(* Logix 5000 project; controller NWGG_Treater_Dayton vendor 1 type 14 code 238 rev 35.11; software revision 35.00; part 2 of 5 *)

ADD_ON_INSTRUCTION SAI_CheckAlive   (* revision 1.0, vendor Jimmy Gao *)
VAR_INPUT
   HeartBeat : BOOL; {required}
END_VAR
VAR_OUTPUT
   Alive : BOOL; {access Read Only, visible}
END_VAR
VAR
   bResetTimer : BOOL; {access None}
   ons : DINT; {access None}
   TON : TIMER; {access None}
END_VAR

ROUTINE Logic   (* ladder *)
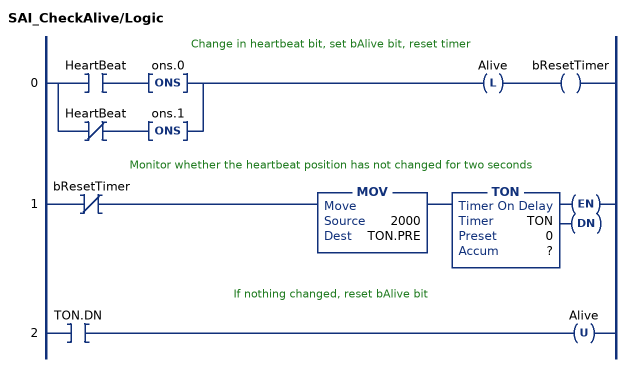
   // Change in heartbeat bit, set bAlive bit, reset timer
   0: [XIC(HeartBeat) ONS(ons.0) ,XIO(HeartBeat) ONS(ons.1) ]OTL(Alive)OTE(bResetTimer);
   // Monitor whether the heartbeat position has not changed for two seconds
   1: XIO(bResetTimer)MOV(2000,TON.PRE)TON(TON,?,?);
   // If nothing changed, reset bAlive bit
   2: XIC(TON.DN)OTU(Alive);
END_ROUTINE
END_ADD_ON_INSTRUCTION

ADD_ON_INSTRUCTION SAI_IND_CalFree   (* revision 1.0, vendor Griffin Hodnett *)
VAR_INPUT
   RatedCapacity : REAL; {required}
   ScaleUnit : DINT; {required}
   RatedOutput : REAL; {access None, required}
   Start : BOOL; {visible}
END_VAR
VAR_OUTPUT
   Done : BOOL; {access Read Only, visible}
   Error : BOOL; {access Read Only, visible}
   Status : DINT; {access Read Only, visible}
END_VAR
VAR_IN_OUT
   MSG_CalFreeTrigger : MESSAGE; {required}
   MSG_CalFreeStatus : MESSAGE; {required}
   MSG_CalFreeUnit : MESSAGE; {required}
   MSG_CalFreeCellCapacity : MESSAGE; {required}
   MSG_CalFreeCellOutput : MESSAGE; {required}
   TmpTrigger : INT; {required}
   TmpAdjStatus : INT; {required}
END_VAR
VAR
   ons : DINT; {access None}
   Step : INT; {access None}
   TON : TIMER[7]; {access None}
   EnterAdj : BOOL; {access None}
   EnterCancel : BOOL; {access None}
END_VAR

ROUTINE Logic   (* ladder *)
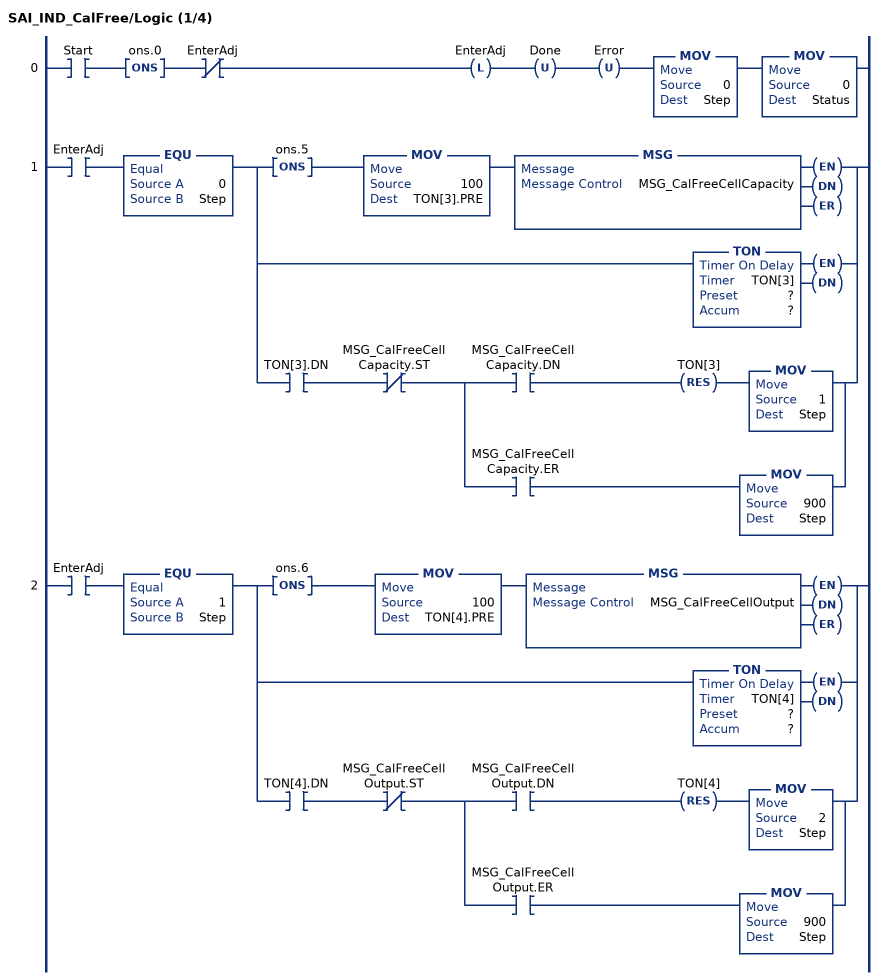
   0: XIC(Start)ONS(ons.0)XIO(EnterAdj)OTL(EnterAdj)OTU(Done)OTU(Error)MOV(0,Step)MOV(0,Status);
   1: XIC(EnterAdj)EQU(0,Step)[[ONS(ons.5) MOV(100,TON[3].PRE) MSG(MSG_CalFreeCellCapacity) ,TON(TON[3],?,?) ] ,XIC(TON[3].DN) XIO(MSG_CalFreeCellCapacity.ST) [XIC(MSG_CalFreeCellCapacity.DN) RES(TON[3]) MOV(1,Step) ,XIC(MSG_CalFreeCellCapacity.ER) MOV(900,Step) ] ];
   2: XIC(EnterAdj)EQU(1,Step)[[ONS(ons.6) MOV(100,TON[4].PRE) MSG(MSG_CalFreeCellOutput) ,TON(TON[4],?,?) ] ,XIC(TON[4].DN) XIO(MSG_CalFreeCellOutput.ST) [XIC(MSG_CalFreeCellOutput.DN) RES(TON[4]) MOV(2,Step) ,XIC(MSG_CalFreeCellOutput.ER) MOV(900,Step) ] ];
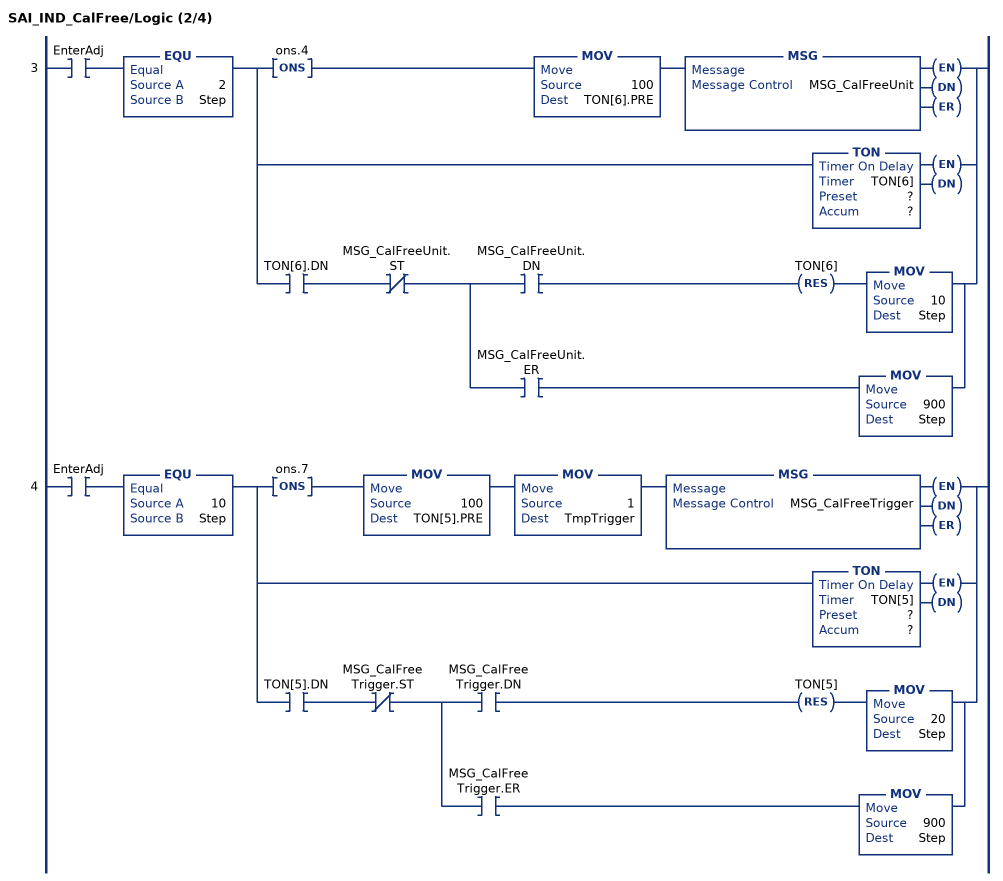
   3: XIC(EnterAdj)EQU(2,Step)[[ONS(ons.4) MOV(100,TON[6].PRE) MSG(MSG_CalFreeUnit) ,TON(TON[6],?,?) ] ,XIC(TON[6].DN) XIO(MSG_CalFreeUnit.ST) [XIC(MSG_CalFreeUnit.DN) RES(TON[6]) MOV(10,Step) ,XIC(MSG_CalFreeUnit.ER) MOV(900,Step) ] ];
   4: XIC(EnterAdj)EQU(10,Step)[[ONS(ons.7) MOV(100,TON[5].PRE) MOV(1,TmpTrigger) MSG(MSG_CalFreeTrigger) ,TON(TON[5],?,?) ] ,XIC(TON[5].DN) XIO(MSG_CalFreeTrigger.ST) [XIC(MSG_CalFreeTrigger.DN) RES(TON[5]) MOV(20,Step) ,XIC(MSG_CalFreeTrigger.ER) MOV(900,Step) ] ];
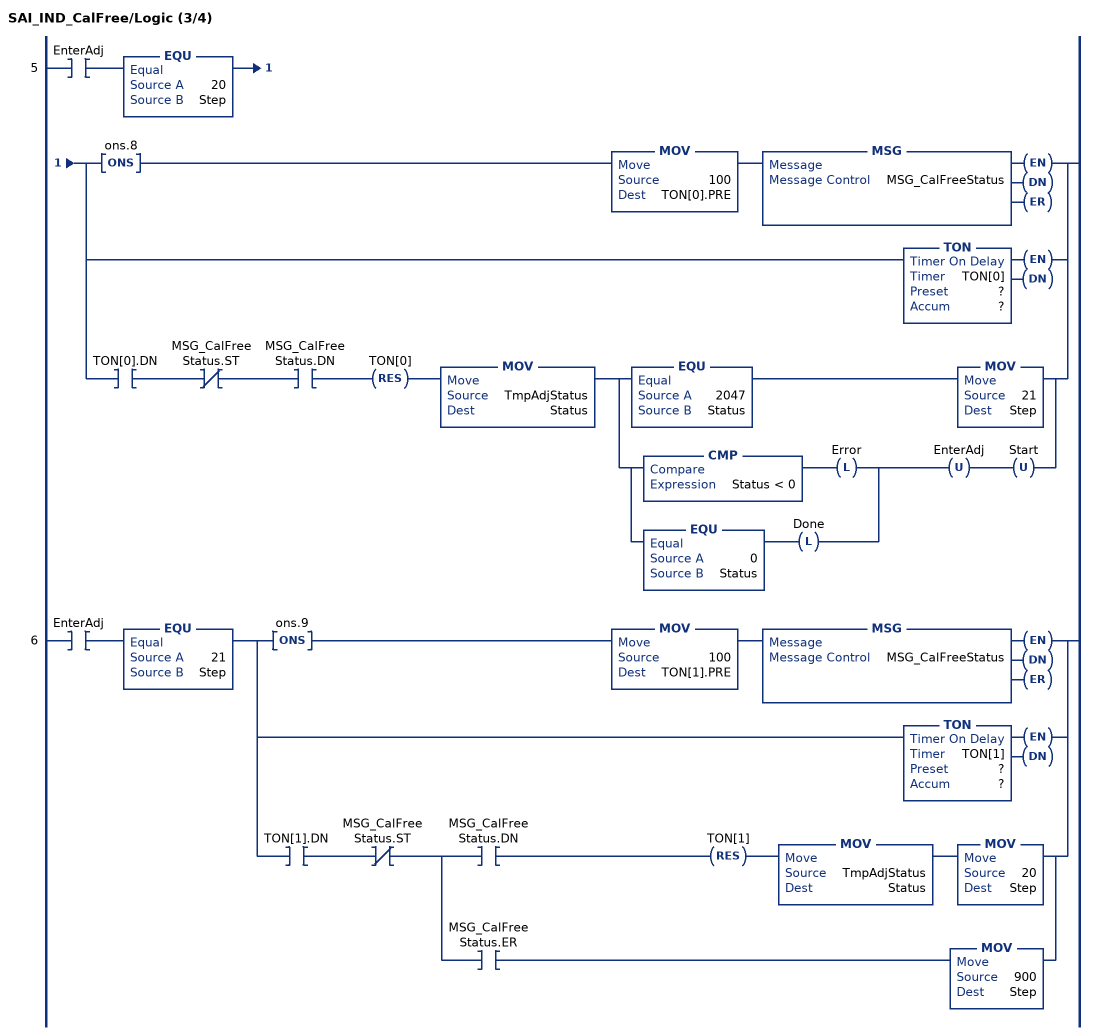
   5: XIC(EnterAdj)EQU(20,Step)[[ONS(ons.8) MOV(100,TON[0].PRE) MSG(MSG_CalFreeStatus) ,TON(TON[0],?,?) ] ,XIC(TON[0].DN) XIO(MSG_CalFreeStatus.ST) XIC(MSG_CalFreeStatus.DN) RES(TON[0]) MOV(TmpAdjStatus,Status) [EQU(2047,Status) MOV(21,Step) ,[CMP(Status < 0) OTL(Error) ,EQU(0,Status) OTL(Done) ] OTU(EnterAdj) OTU(Start) ] ];
   6: XIC(EnterAdj)EQU(21,Step)[[ONS(ons.9) MOV(100,TON[1].PRE) MSG(MSG_CalFreeStatus) ,TON(TON[1],?,?) ] ,XIC(TON[1].DN) XIO(MSG_CalFreeStatus.ST) [XIC(MSG_CalFreeStatus.DN) RES(TON[1]) MOV(TmpAdjStatus,Status) MOV(20,Step) ,XIC(MSG_CalFreeStatus.ER) MOV(900,Step) ] ];
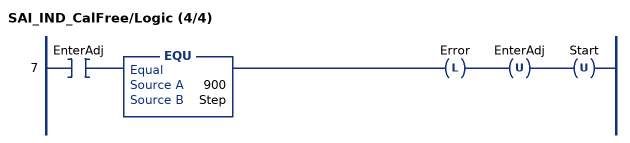
   7: XIC(EnterAdj)EQU(900,Step)OTL(Error)OTU(EnterAdj)OTU(Start);
END_ROUTINE
END_ADD_ON_INSTRUCTION

ADD_ON_INSTRUCTION SAI_IND_ReadAdjustSettings   (* revision 1.0, vendor Griffin Hodnett *)
VAR_INPUT
   Read : BOOL; {visible}
END_VAR
VAR_OUTPUT
   ScaleCapacity : REAL; {visible}
   Increment : REAL; {visible}
   Done : BOOL; {access Read Only, visible}
   Error : BOOL; {access Read Only, visible}
END_VAR
VAR_IN_OUT
   MSG_ReadCap : MESSAGE; {required}
   MSG_ReadInc : MESSAGE; {required}
   TmpInc : REAL; {required}
   TmpCapacity : REAL; {required}
END_VAR
VAR
   TON : TIMER[1]; {access None}
   Step : INT; {access None}
   Get_Values : BOOL; {access None}
   ons : DINT; {access None}
END_VAR

ROUTINE Logic   (* ladder *)
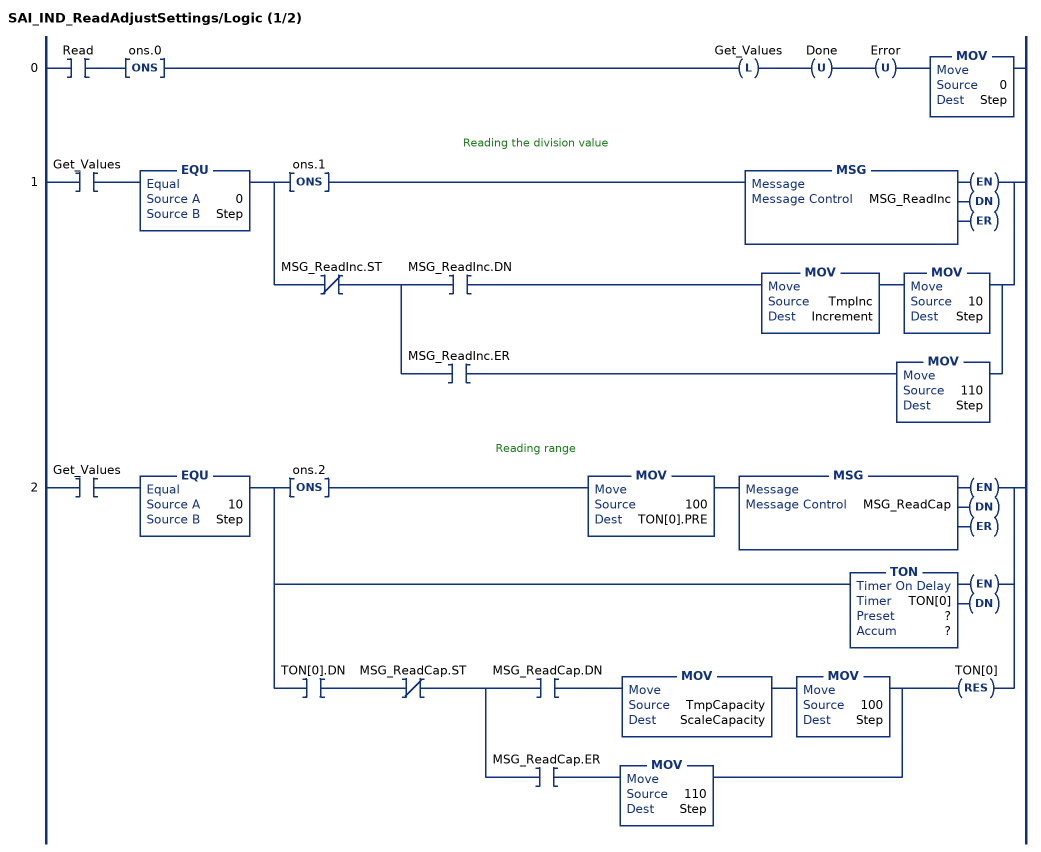
   0: XIC(Read)ONS(ons.0)OTL(Get_Values)OTU(Done)OTU(Error)MOV(0,Step);
   // Reading the division value
   1: XIC(Get_Values)EQU(0,Step)[ONS(ons.1) MSG(MSG_ReadInc) ,XIO(MSG_ReadInc.ST) [XIC(MSG_ReadInc.DN) MOV(TmpInc,Increment) MOV(10,Step) ,XIC(MSG_ReadInc.ER) MOV(110,Step) ] ];
   // Reading range
   2: XIC(Get_Values)EQU(10,Step)[[ONS(ons.2) MOV(100,TON[0].PRE) MSG(MSG_ReadCap) ,TON(TON[0],?,?) ] ,XIC(TON[0].DN) XIO(MSG_ReadCap.ST) [XIC(MSG_ReadCap.DN) MOV(TmpCapacity,ScaleCapacity) MOV(100,Step) ,XIC(MSG_ReadCap.ER) MOV(110,Step) ] RES(TON[0]) ];
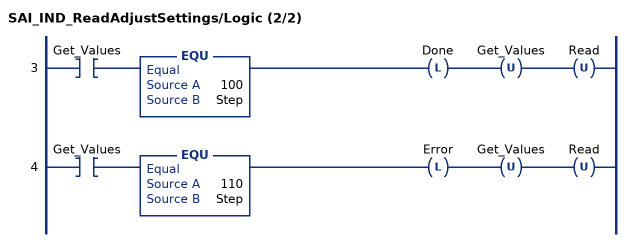
   3: XIC(Get_Values)EQU(100,Step)OTL(Done)OTU(Get_Values)OTU(Read);
   4: XIC(Get_Values)EQU(110,Step)OTL(Error)OTU(Get_Values)OTU(Read);
END_ROUTINE
END_ADD_ON_INSTRUCTION

ADD_ON_INSTRUCTION SAI_IND_SpanAdjust   (* revision 1.0, vendor Griffin Hodnett *)
VAR_INPUT
   LinearityRange : INT; {access None, required}
   Hi_Weight : REAL; {visible}
   Mid_Weight : REAL; {visible}
   Low_Weight : REAL; {visible}
   xLow_Weight : REAL; {visible}
   Start : BOOL; {visible}
END_VAR
VAR_OUTPUT
   CurrentWeight : REAL; {access Read Only, visible}
END_VAR
VAR_INPUT
   ConfirmWeight : BOOL; {visible}
   Cancel : BOOL; {visible}
END_VAR
VAR_OUTPUT
   Done : BOOL; {access Read Only, visible}
   Error : BOOL; {access Read Only, visible}
   Cancelled : BOOL; {access Read Only, visible}
   LoadWeight : BOOL; {access Read Only, visible}
END_VAR
VAR_INPUT
   DataOK : BOOL; {required}
END_VAR
VAR_OUTPUT
   Status : INT; {access Read Only, visible}
   CurrentPoint : DINT; {access Read Only, visible}
END_VAR
VAR_IN_OUT
   MSG_CancelAdj : MESSAGE; {required}
   MSG_StartSpanAdj : MESSAGE; {required}
   MSG_LinearityRange : MESSAGE; {required}
   MSG_ReadAdjStatus : MESSAGE; {required}
   MSG_ValidateAdj : MESSAGE; {required}
   TmpTrigger : SINT; {required}
   TmpAdjStatus : INT; {required}
   TmpSpanAdjWeight : REAL; {required}
END_VAR
VAR
   Step : INT; {access None}
   TON : TIMER[3]; {access None}
   ons : DINT; {access None}
   EnterCancel : BOOL; {access None}
   EnterAdj : BOOL; {access None}
   WeightCheck : BOOL; {access None}
END_VAR

ROUTINE Logic   (* ladder *)
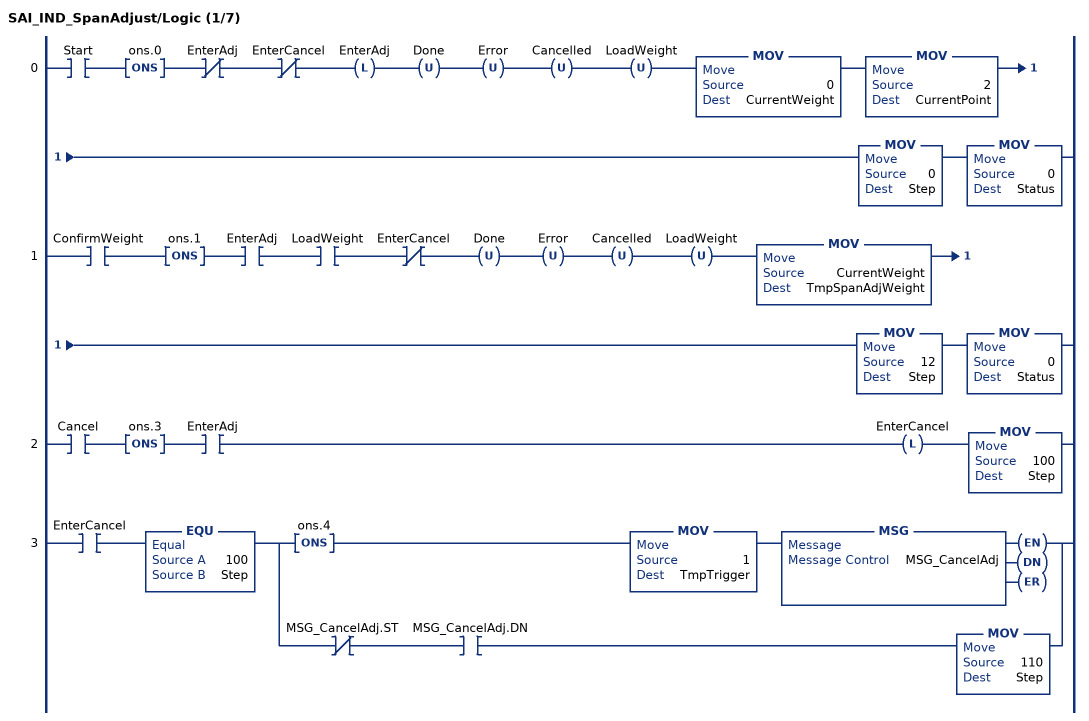
   0: XIC(Start)ONS(ons.0)XIO(EnterAdj)XIO(EnterCancel)OTL(EnterAdj)OTU(Done)OTU(Error)OTU(Cancelled)OTU(LoadWeight)MOV(0,CurrentWeight)MOV(2,CurrentPoint)MOV(0,Step)MOV(0,Status);
   1: XIC(ConfirmWeight)ONS(ons.1)XIC(EnterAdj)XIC(LoadWeight)XIO(EnterCancel)OTU(Done)OTU(Error)OTU(Cancelled)OTU(LoadWeight)MOV(CurrentWeight,TmpSpanAdjWeight)MOV(12,Step)MOV(0,Status);
   2: XIC(Cancel)ONS(ons.3)XIC(EnterAdj)OTL(EnterCancel)MOV(100,Step);
   3: XIC(EnterCancel)EQU(100,Step)[ONS(ons.4) MOV(1,TmpTrigger) MSG(MSG_CancelAdj) ,XIO(MSG_CancelAdj.ST) XIC(MSG_CancelAdj.DN) MOV(110,Step) ];
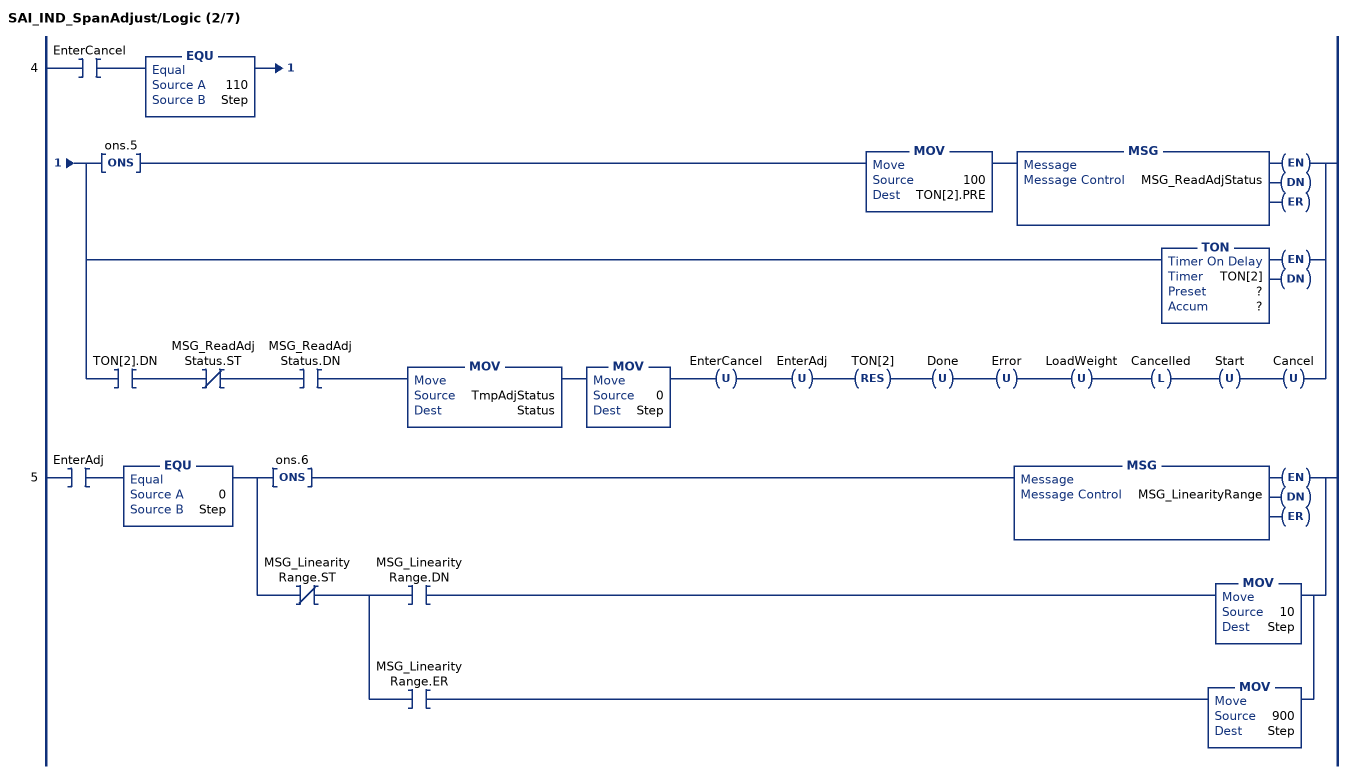
   4: XIC(EnterCancel)EQU(110,Step)[[ONS(ons.5) MOV(100,TON[2].PRE) MSG(MSG_ReadAdjStatus) ,TON(TON[2],?,?) ] ,XIC(TON[2].DN) XIO(MSG_ReadAdjStatus.ST) XIC(MSG_ReadAdjStatus.DN) MOV(TmpAdjStatus,Status) MOV(0,Step) OTU(EnterCancel) OTU(EnterAdj) RES(TON[2]) OTU(Done) OTU(Error) OTU(LoadWeight) OTL(Cancelled) OTU(Start) OTU(Cancel) ];
   5: XIC(EnterAdj)EQU(0,Step)[ONS(ons.6) MSG(MSG_LinearityRange) ,XIO(MSG_LinearityRange.ST) [XIC(MSG_LinearityRange.DN) MOV(10,Step) ,XIC(MSG_LinearityRange.ER) MOV(900,Step) ] ];
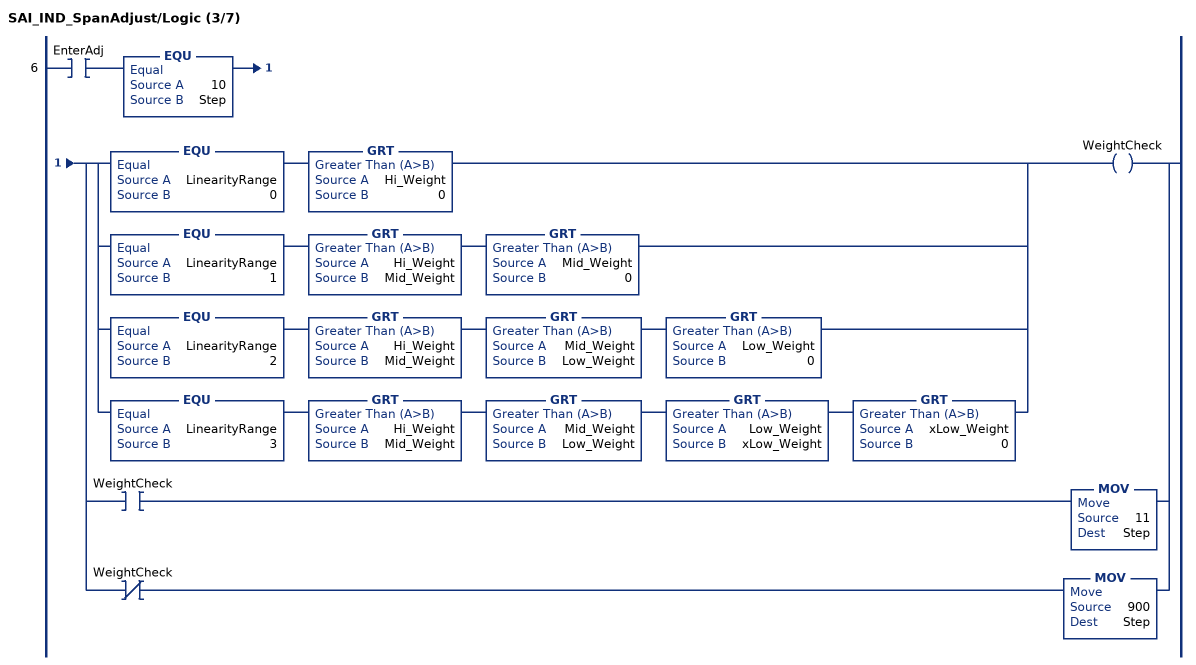
   6: XIC(EnterAdj)EQU(10,Step)[[EQU(LinearityRange,0) GRT(Hi_Weight,0) ,[EQU(LinearityRange,1) GRT(Hi_Weight,Mid_Weight) GRT(Mid_Weight,0) ,[EQU(LinearityRange,2) GRT(Hi_Weight,Mid_Weight) GRT(Mid_Weight,Low_Weight) GRT(Low_Weight,0) ,EQU(LinearityRange,3) GRT(Hi_Weight,Mid_Weight) GRT(Mid_Weight,Low_Weight) GRT(Low_Weight,xLow_Weight) GRT(xLow_Weight,0) ] ] ] OTE(WeightCheck) ,[XIC(WeightCheck) MOV(11,Step) ,XIO(WeightCheck) MOV(900,Step) ] ];
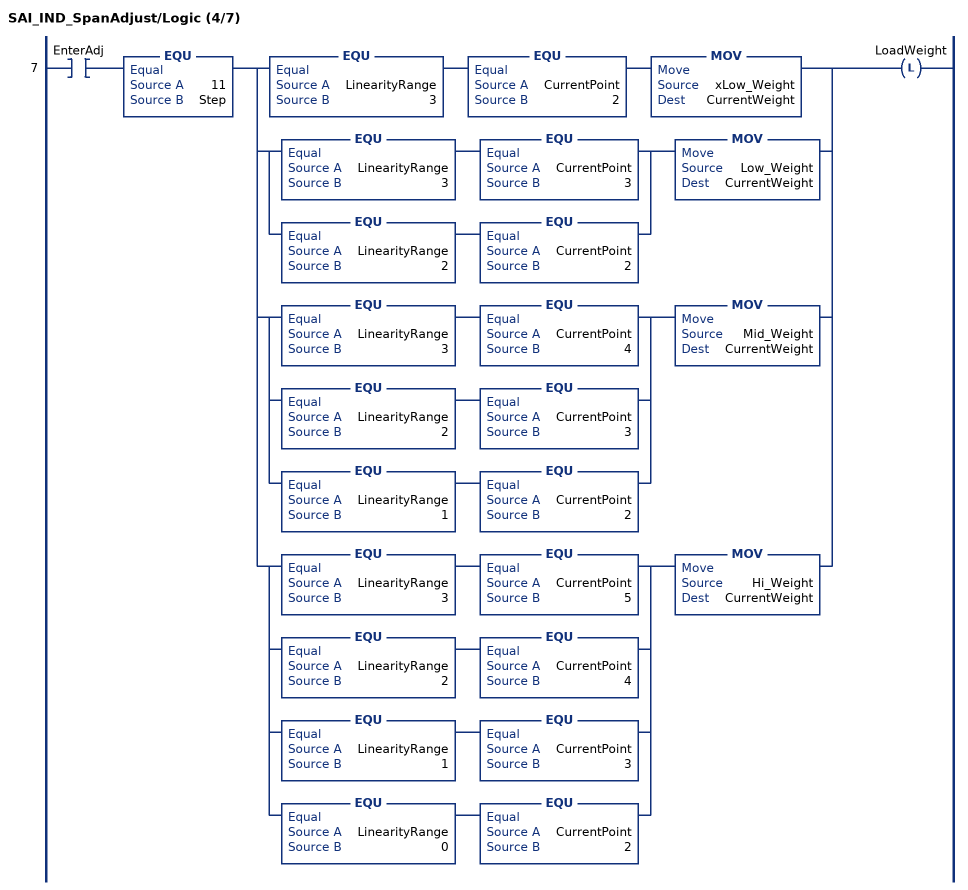
   7: XIC(EnterAdj)EQU(11,Step)[EQU(LinearityRange,3) EQU(CurrentPoint,2) MOV(xLow_Weight,CurrentWeight) ,[[[EQU(LinearityRange,3) EQU(CurrentPoint,3) ,EQU(LinearityRange,2) EQU(CurrentPoint,2) ] MOV(Low_Weight,CurrentWeight) ,[EQU(LinearityRange,3) EQU(CurrentPoint,4) ,[EQU(LinearityRange,2) EQU(CurrentPoint,3) ,EQU(LinearityRange,1) EQU(CurrentPoint,2) ] ] MOV(Mid_Weight,CurrentWeight) ] ,[EQU(LinearityRange,3) EQU(CurrentPoint,5) ,[EQU(LinearityRange,2) EQU(CurrentPoint,4) ,[EQU(LinearityRange,1) EQU(CurrentPoint,3) ,EQU(LinearityRange,0) EQU(CurrentPoint,2) ] ] ] MOV(Hi_Weight,CurrentWeight) ] ]OTL(LoadWeight);
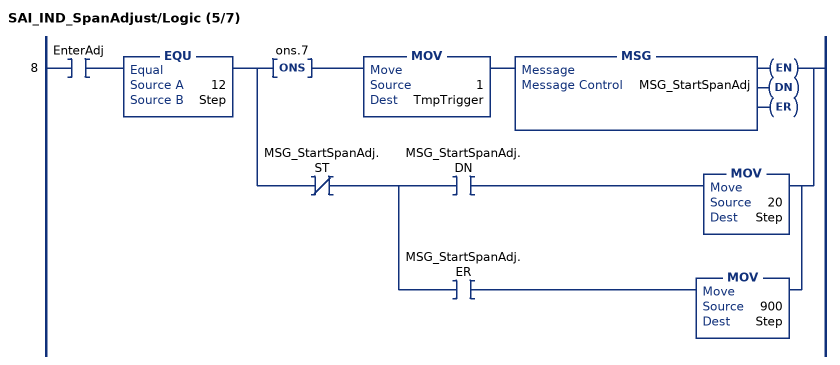
   8: XIC(EnterAdj)EQU(12,Step)[ONS(ons.7) MOV(1,TmpTrigger) MSG(MSG_StartSpanAdj) ,XIO(MSG_StartSpanAdj.ST) [XIC(MSG_StartSpanAdj.DN) MOV(20,Step) ,XIC(MSG_StartSpanAdj.ER) MOV(900,Step) ] ];
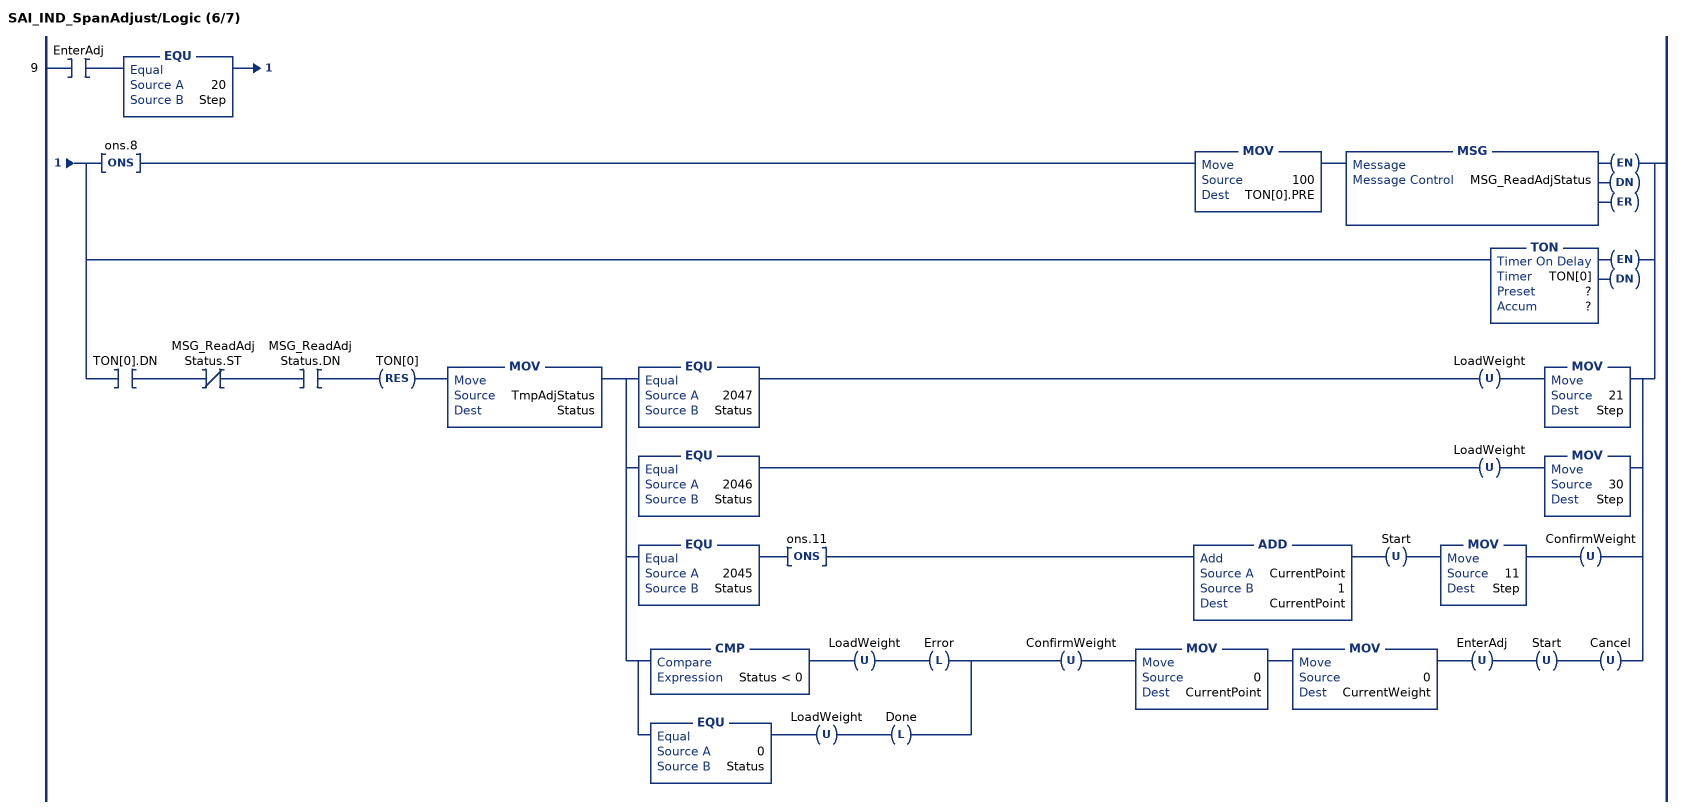
   9: XIC(EnterAdj)EQU(20,Step)[[ONS(ons.8) MOV(100,TON[0].PRE) MSG(MSG_ReadAdjStatus) ,TON(TON[0],?,?) ] ,XIC(TON[0].DN) XIO(MSG_ReadAdjStatus.ST) XIC(MSG_ReadAdjStatus.DN) RES(TON[0]) MOV(TmpAdjStatus,Status) [EQU(2047,Status) OTU(LoadWeight) MOV(21,Step) ,[[EQU(2046,Status) OTU(LoadWeight) MOV(30,Step) ,EQU(2045,Status) ONS(ons.11) ADD(CurrentPoint,1,CurrentPoint) OTU(Start) MOV(11,Step) OTU(ConfirmWeight) ] ,[CMP(Status < 0) OTU(LoadWeight) OTL(Error) ,EQU(0,Status) OTU(LoadWeight) OTL(Done) ] OTU(ConfirmWeight) MOV(0,CurrentPoint) MOV(0,CurrentWeight) OTU(EnterAdj) OTU(Start) OTU(Cancel) ] ] ];
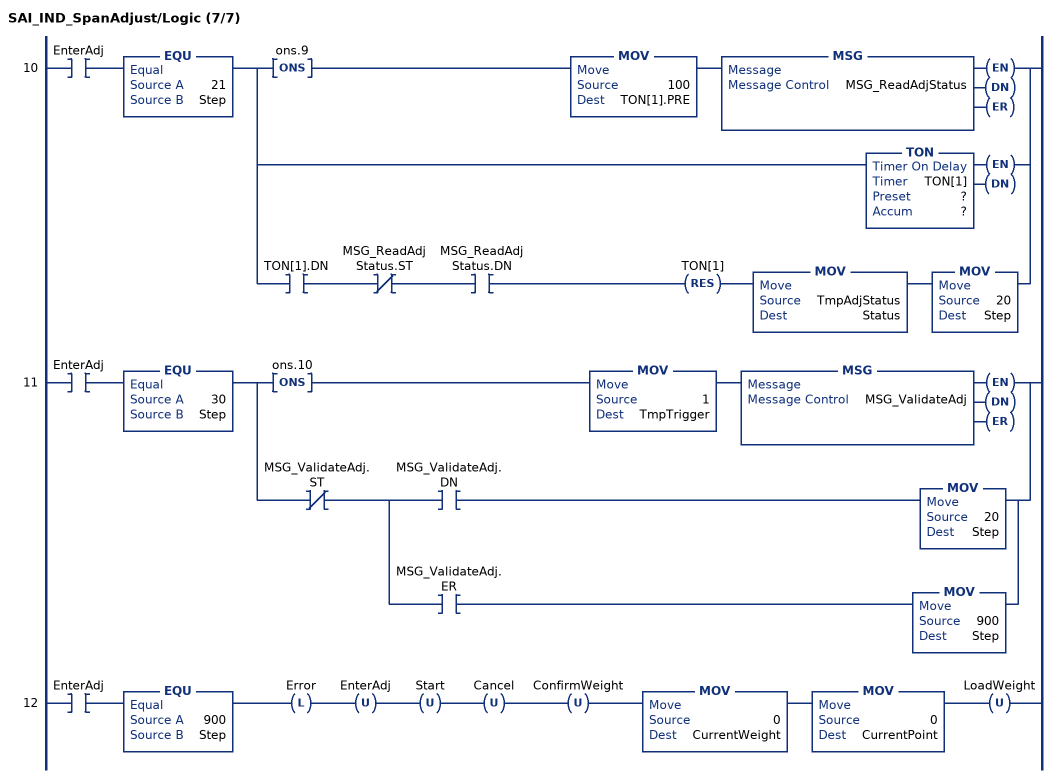
   10: XIC(EnterAdj)EQU(21,Step)[[ONS(ons.9) MOV(100,TON[1].PRE) MSG(MSG_ReadAdjStatus) ,TON(TON[1],?,?) ] ,XIC(TON[1].DN) XIO(MSG_ReadAdjStatus.ST) XIC(MSG_ReadAdjStatus.DN) RES(TON[1]) MOV(TmpAdjStatus,Status) MOV(20,Step) ];
   11: XIC(EnterAdj)EQU(30,Step)[ONS(ons.10) MOV(1,TmpTrigger) MSG(MSG_ValidateAdj) ,XIO(MSG_ValidateAdj.ST) [XIC(MSG_ValidateAdj.DN) MOV(20,Step) ,XIC(MSG_ValidateAdj.ER) MOV(900,Step) ] ];
   12: XIC(EnterAdj)EQU(900,Step)OTL(Error)OTU(EnterAdj)OTU(Start)OTU(Cancel)OTU(ConfirmWeight)MOV(0,CurrentWeight)MOV(0,CurrentPoint)OTU(LoadWeight);
END_ROUTINE
END_ADD_ON_INSTRUCTION

ADD_ON_INSTRUCTION SAI_IND_WeightProc   (* revision 1.0, vendor Griffin Hodnett *)
VAR_INPUT
   WeightCmd : INT; {visible}
   TareImmediate : BOOL; {visible}
   TareStable : BOOL; {visible}
   ZeroImmediate : BOOL; {visible}
   ZeroStable : BOOL; {visible}
   PreTareValue : REAL; {visible}
   PreTare : BOOL; {visible}
   ClearTare : BOOL; {visible}
   MB_Value : REAL; {access Read Only, required}
   MB_Response : INT; {access Read Only, required}
END_VAR
VAR_IN_OUT
   MB_CmdValue : REAL; {required}
END_VAR
VAR_OUTPUT
   MB_Command : INT; {access Read Only, required}
END_VAR
VAR_INPUT
   DataOK : BOOL; {access Read Only, required}
   Motion : BOOL; {access Read Only, required}
   NetMode : BOOL; {required}
   Alarm : BOOL; {required}
END_VAR
VAR_OUTPUT
   RealTimeWeight : REAL; {access Read Only, visible}
   StableWeight : REAL; {access Read Only, visible}
   Done : BOOL; {access Read Only, visible}
   Error : BOOL; {access Read Only, visible}
END_VAR
VAR
   WriteTrigger : BOOL; {access None}
   RestoreTrigger : BOOL; {access None}
   Command : INT; {access None}
   ons : DINT; {access None}
   Prev_WeightCmd : DINT; {access None}
END_VAR

ROUTINE Logic   (* ladder *)
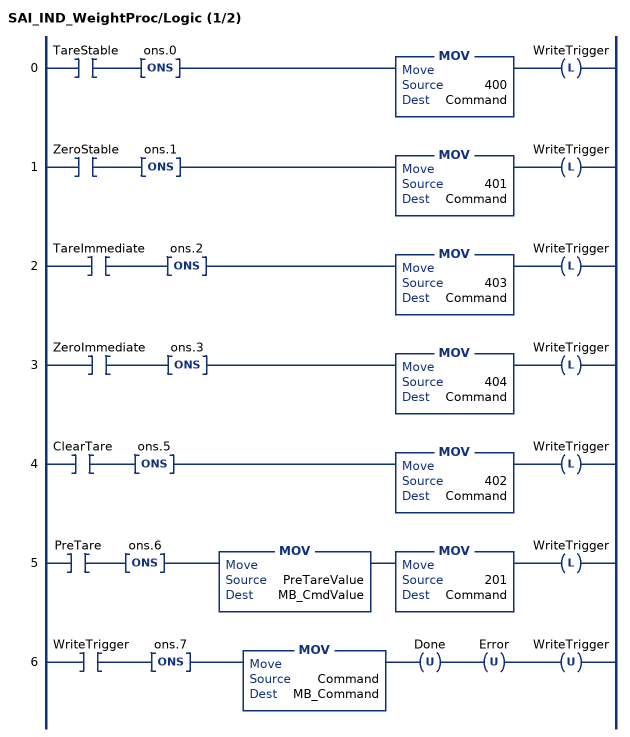
   0: XIC(TareStable)ONS(ons.0)MOV(400,Command)OTL(WriteTrigger);
   1: XIC(ZeroStable)ONS(ons.1)MOV(401,Command)OTL(WriteTrigger);
   2: XIC(TareImmediate)ONS(ons.2)MOV(403,Command)OTL(WriteTrigger);
   3: XIC(ZeroImmediate)ONS(ons.3)MOV(404,Command)OTL(WriteTrigger);
   4: XIC(ClearTare)ONS(ons.5)MOV(402,Command)OTL(WriteTrigger);
   5: XIC(PreTare)ONS(ons.6)MOV(PreTareValue,MB_CmdValue)MOV(201,Command)OTL(WriteTrigger);
   6: XIC(WriteTrigger)ONS(ons.7)MOV(Command,MB_Command)OTU(Done)OTU(Error)OTU(WriteTrigger);
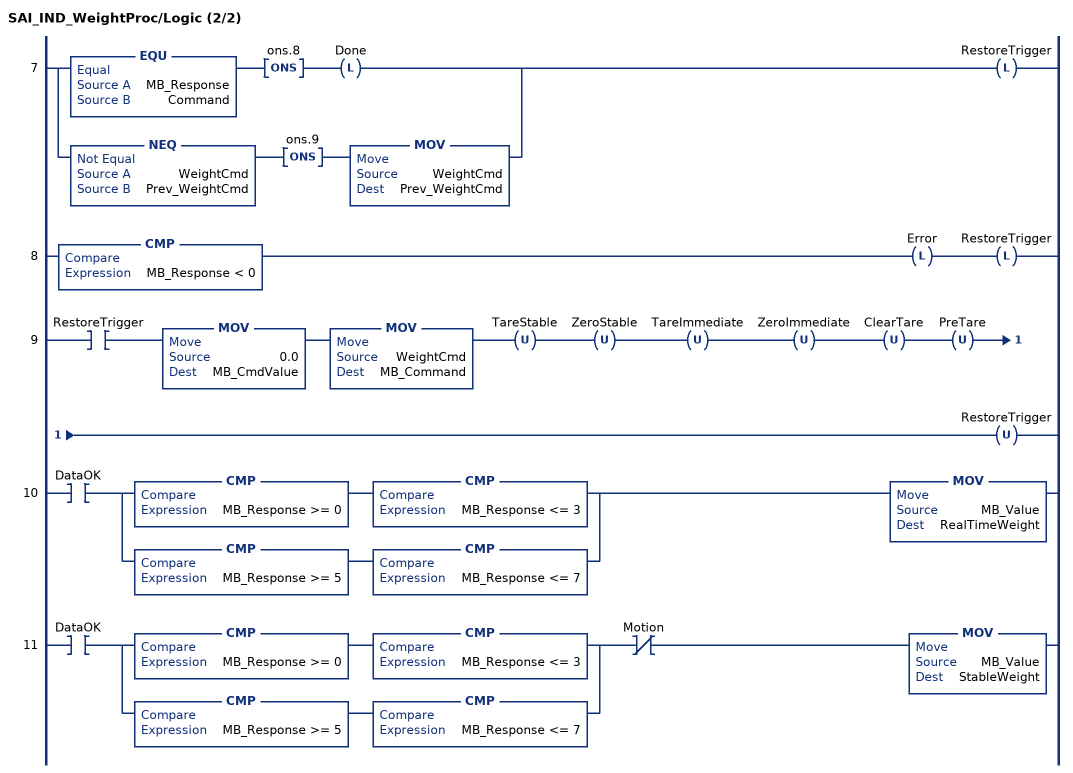
   7: [EQU(MB_Response,Command) ONS(ons.8) OTL(Done) ,NEQ(WeightCmd,Prev_WeightCmd) ONS(ons.9) MOV(WeightCmd,Prev_WeightCmd) ]OTL(RestoreTrigger);
   8: CMP(MB_Response < 0)OTL(Error)OTL(RestoreTrigger);
   9: XIC(RestoreTrigger)MOV(0.0,MB_CmdValue)MOV(WeightCmd,MB_Command)OTU(TareStable)OTU(ZeroStable)OTU(TareImmediate)OTU(ZeroImmediate)OTU(ClearTare)OTU(PreTare)OTU(RestoreTrigger);
   10: XIC(DataOK)[CMP(MB_Response >= 0) CMP(MB_Response <= 3) ,CMP(MB_Response >= 5) CMP(MB_Response <= 7) ]MOV(MB_Value,RealTimeWeight);
   11: XIC(DataOK)[CMP(MB_Response >= 0) CMP(MB_Response <= 3) ,CMP(MB_Response >= 5) CMP(MB_Response <= 7) ]XIO(Motion)MOV(MB_Value,StableWeight);
END_ROUTINE
END_ADD_ON_INSTRUCTION

ADD_ON_INSTRUCTION SAI_IND_WriteAdjustSettings   (* revision 1.0, vendor Griffin Hodnett *)
VAR_INPUT
   ScaleCapacity : REAL; {required}
   Increment : REAL; {required}
   Write : BOOL; {visible}
END_VAR
VAR_OUTPUT
   Done : BOOL; {access Read Only, visible}
   Error : BOOL; {access Read Only, visible}
END_VAR
VAR_IN_OUT
   MSG_WriteCap : MESSAGE; {required}
   MSG_WriteInc : MESSAGE; {required}
END_VAR
VAR
   ons : DINT; {access None}
   Step : INT; {access None}
   TON : TIMER[2]; {access None}
   Write_Values : BOOL; {access None}
END_VAR

ROUTINE Logic   (* ladder *)
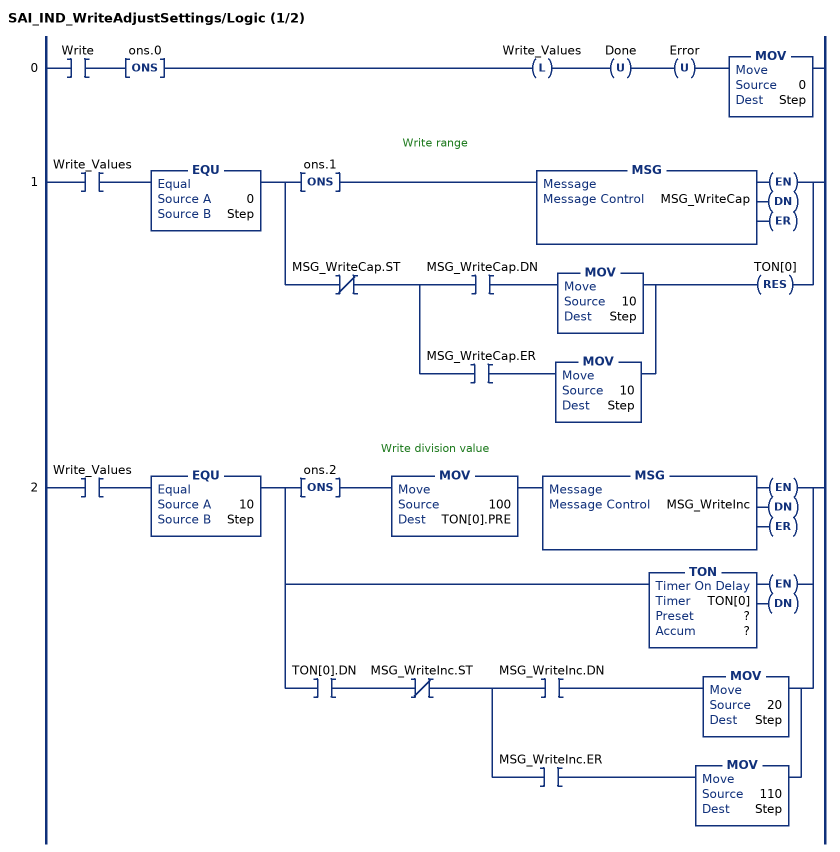
   0: XIC(Write)ONS(ons.0)OTL(Write_Values)OTU(Done)OTU(Error)MOV(0,Step);
   // Write range
   1: XIC(Write_Values)EQU(0,Step)[ONS(ons.1) MSG(MSG_WriteCap) ,XIO(MSG_WriteCap.ST) [XIC(MSG_WriteCap.DN) MOV(10,Step) ,XIC(MSG_WriteCap.ER) MOV(10,Step) ] RES(TON[0]) ];
   // Write division value
   2: XIC(Write_Values)EQU(10,Step)[[ONS(ons.2) MOV(100,TON[0].PRE) MSG(MSG_WriteInc) ,TON(TON[0],?,?) ] ,XIC(TON[0].DN) XIO(MSG_WriteInc.ST) [XIC(MSG_WriteInc.DN) MOV(20,Step) ,XIC(MSG_WriteInc.ER) MOV(110,Step) ] ];
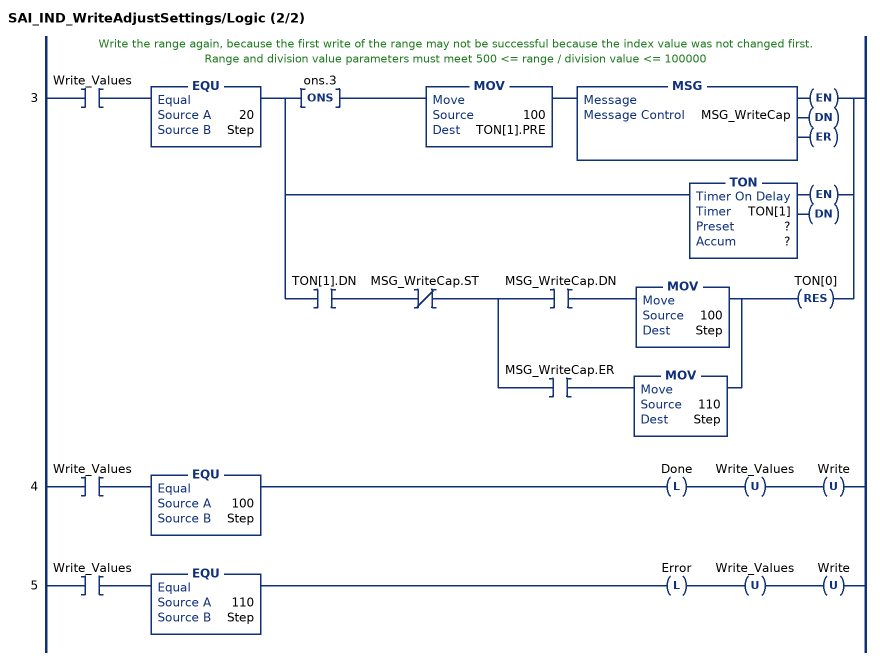
   // Write the range again, because the first write of the range may not be successful because the index value was not changed first.
   // Range and division value parameters must meet 500 <= range / division value <= 100000
   3: XIC(Write_Values)EQU(20,Step)[[ONS(ons.3) MOV(100,TON[1].PRE) MSG(MSG_WriteCap) ,TON(TON[1],?,?) ] ,XIC(TON[1].DN) XIO(MSG_WriteCap.ST) [XIC(MSG_WriteCap.DN) MOV(100,Step) ,XIC(MSG_WriteCap.ER) MOV(110,Step) ] RES(TON[0]) ];
   4: XIC(Write_Values)EQU(100,Step)OTL(Done)OTU(Write_Values)OTU(Write);
   5: XIC(Write_Values)EQU(110,Step)OTL(Error)OTU(Write_Values)OTU(Write);
END_ROUTINE
END_ADD_ON_INSTRUCTION
